// CFC twin of T_SafePulse_UserFB_Tests: the same tests drawn as CFC diagrams, the way a TwinSAFE project is authored.
    FUNCTION_BLOCK T_SafePulse_UserFB_Tests_CFC EXTENDS T_SafeCfcTestSuite
    VAR
    // Test_PulseForDelayTimeWhileInputHeld
    group_1 : T_SafeGroup;
    fb_1 : T_SafePulse_UserFB(group := group_1) := (Parameters := (DelayTime := T#100MS));
    trigStart_1 : R_TRIG;
    t1_1 : TON;
    t2_1 : TON;
    trig1_1 : R_TRIG;
    trig2_1 : R_TRIG;
    // Test_PulseEndsWhenInputDrops
    group_2 : T_SafeGroup;
    fb_2 : T_SafePulse_UserFB(group := group_2) := (Parameters := (DelayTime := T#100MS));
    // Test_StoppedGivesNoOutput
    group_3 : T_SafeGroup;
    fb_3 : T_SafePulse_UserFB(group := group_3) := (Parameters := (DelayTime := T#100MS));
    // Test_InnerBlocksJoinTheGroup
    group_4 : T_SafeGroup;
    fb_4 : T_SafePulse_UserFB(group := group_4);
END_VAR

Test_PulseForDelayTimeWhileInputHeld();
Test_PulseEndsWhenInputDrops();
Test_StoppedGivesNoOutput();
Test_InnerBlocksJoinTheGroup();

METHOD PRIVATE Test_InnerBlocksJoinTheGroup
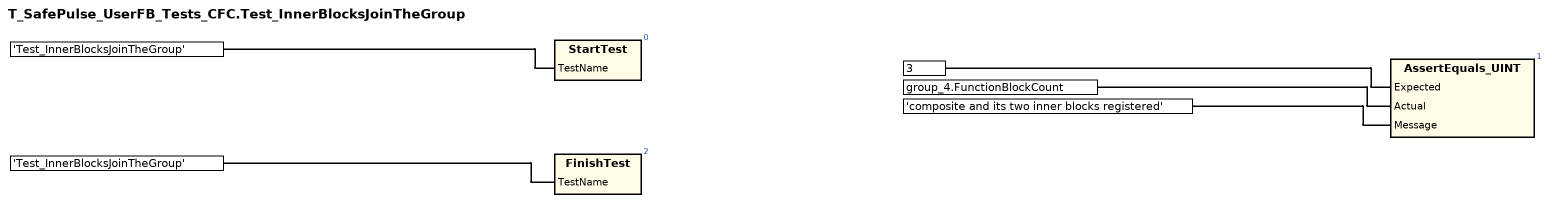
StartTest(TestName := 'Test_InnerBlocksJoinTheGroup');
AssertEquals_UINT(Expected := 3, Actual := group_4.FunctionBlockCount, Message := 'composite and its two inner blocks registered');
FinishTest(TestName := 'Test_InnerBlocksJoinTheGroup');
END_METHOD

METHOD PRIVATE Test_PulseEndsWhenInputDrops
// note: this text did not pass the execution check against the stored diagram
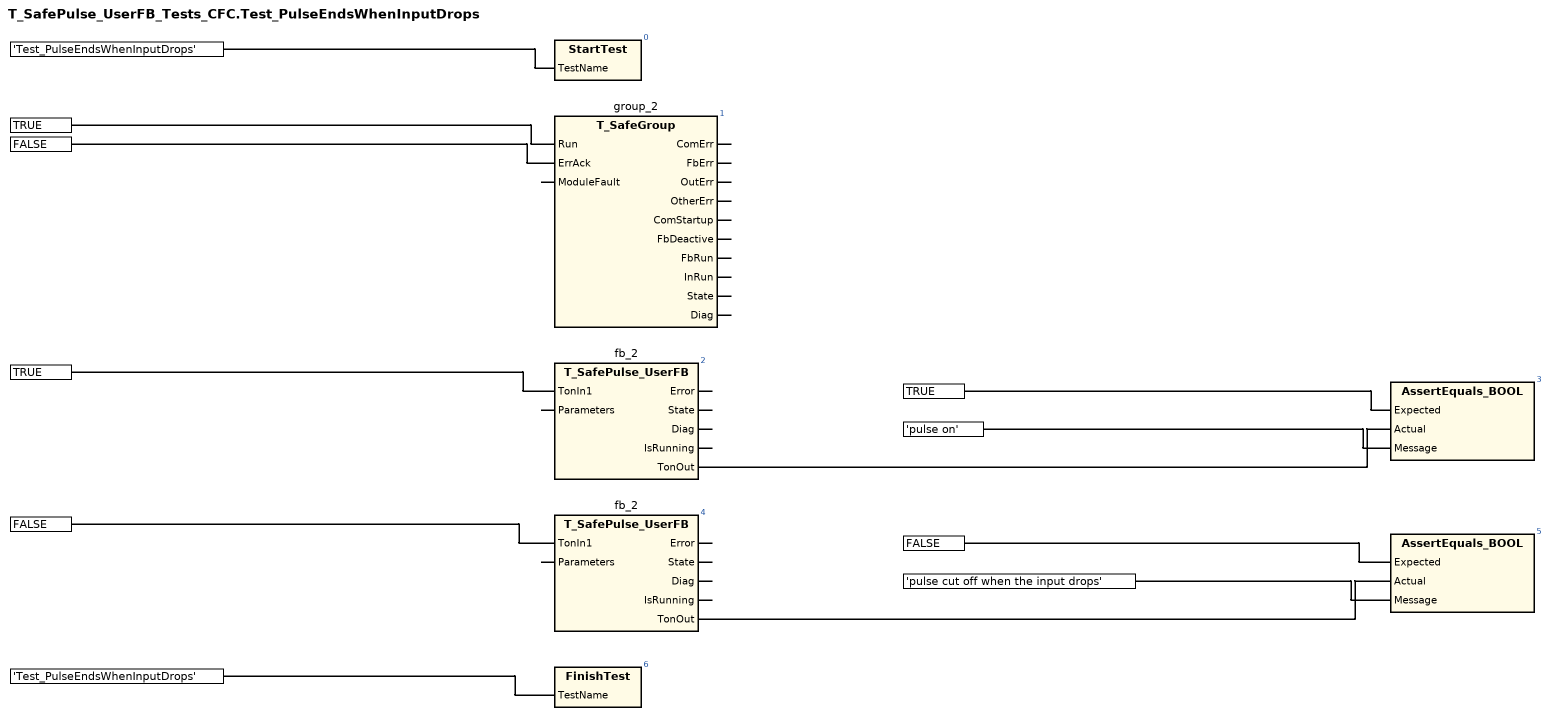
StartTest(TestName := 'Test_PulseEndsWhenInputDrops');
group_2(Run := TRUE, ErrAck := FALSE); // T_SafeGroup
fb_2(TonIn1 := TRUE); // T_SafePulse_UserFB
AssertEquals_BOOL(Expected := TRUE, Actual := fb_2.TonOut, Message := 'pulse on');
fb_2(TonIn1 := FALSE); // T_SafePulse_UserFB
AssertEquals_BOOL(Expected := FALSE, Actual := fb_2.TonOut, Message := 'pulse cut off when the input drops');
FinishTest(TestName := 'Test_PulseEndsWhenInputDrops');
END_METHOD

METHOD PRIVATE Test_PulseForDelayTimeWhileInputHeld
// note: this text did not pass the execution check against the stored diagram
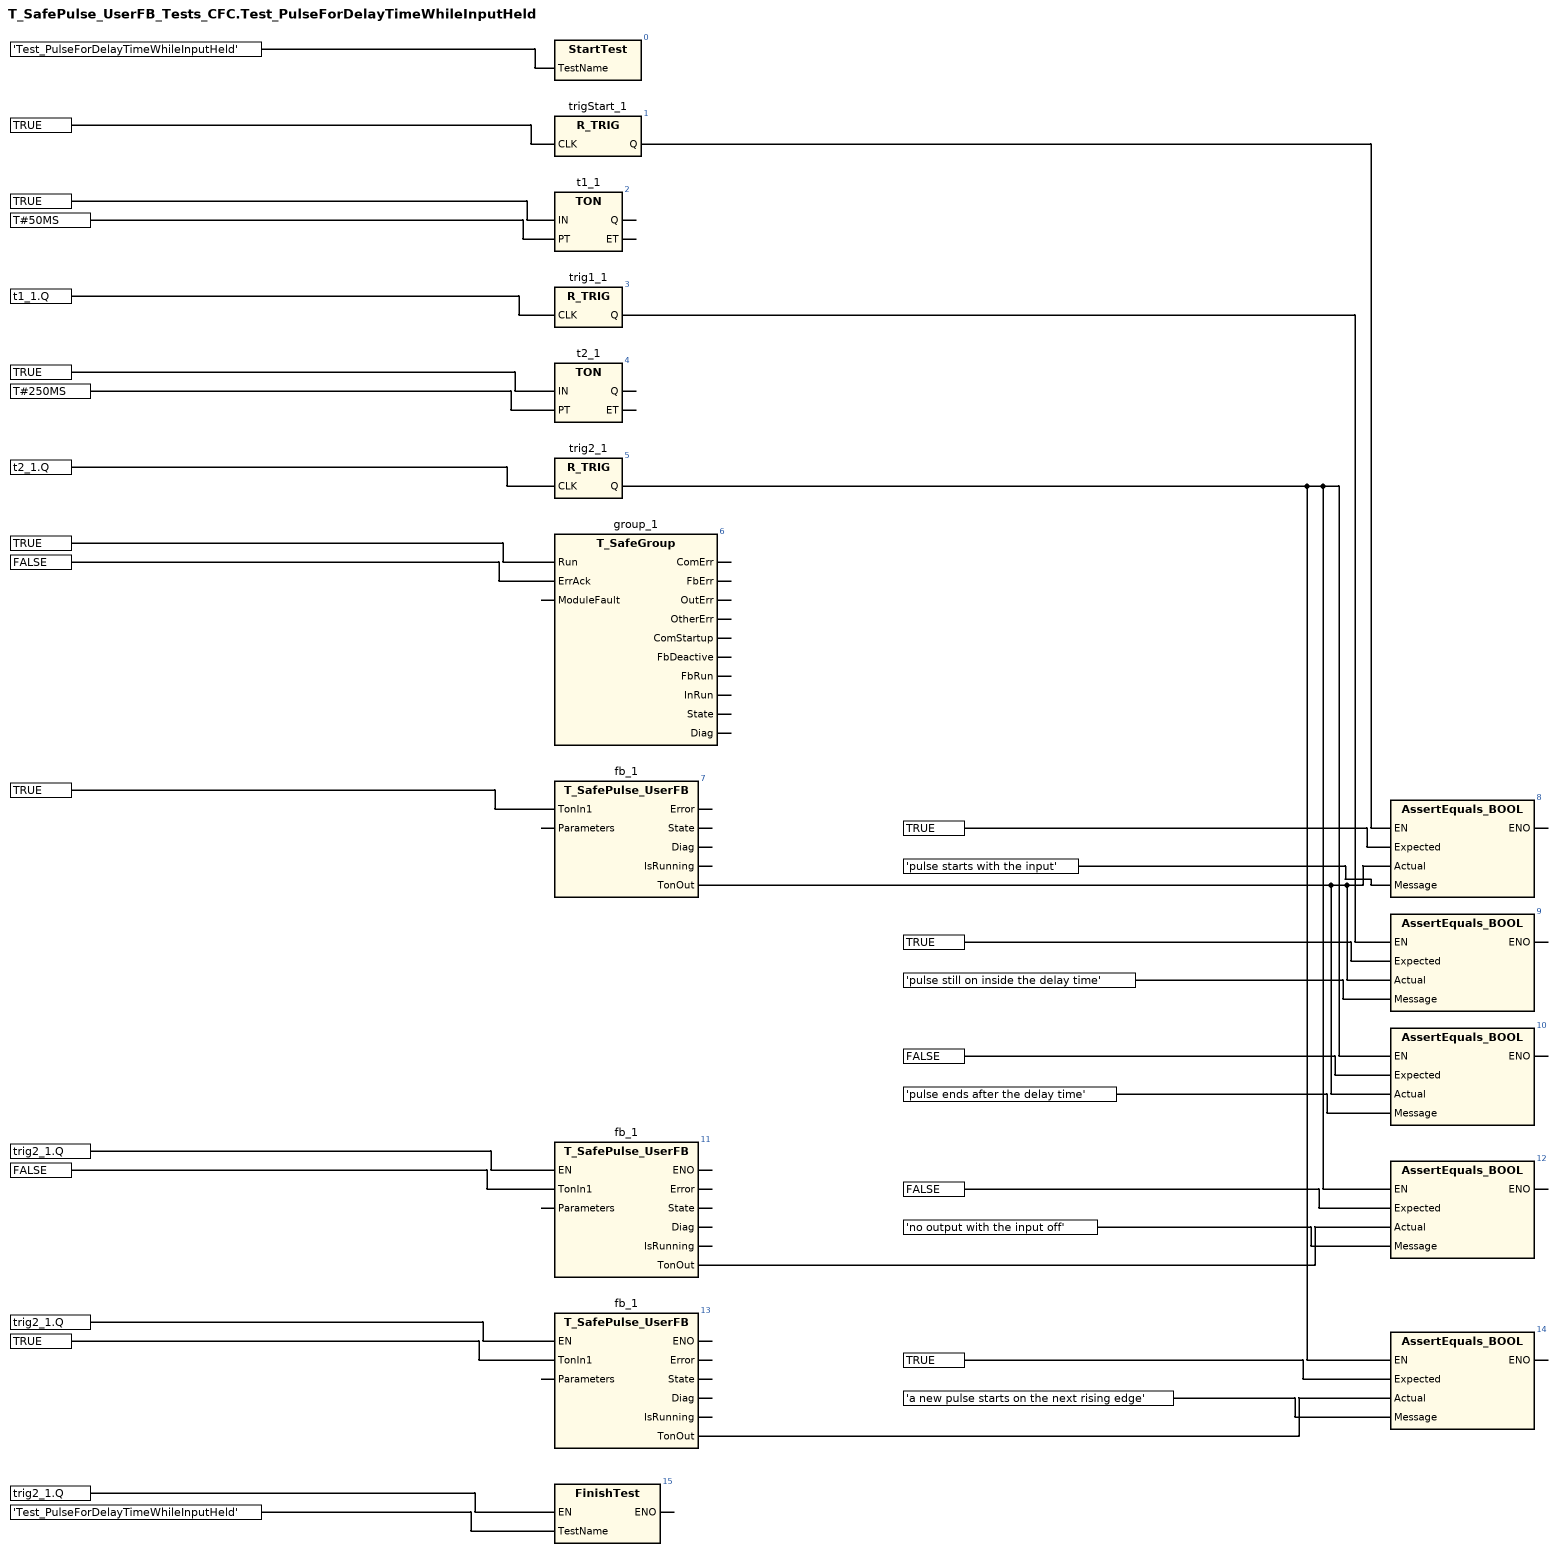
StartTest(TestName := 'Test_PulseForDelayTimeWhileInputHeld');
trigStart_1(CLK := TRUE); // R_TRIG
t1_1(IN := TRUE, PT := T#50MS); // TON
trig1_1(CLK := t1_1.Q); // R_TRIG
t2_1(IN := TRUE, PT := T#250MS); // TON
trig2_1(CLK := t2_1.Q); // R_TRIG
group_1(Run := TRUE, ErrAck := FALSE); // T_SafeGroup
fb_1(TonIn1 := TRUE); // T_SafePulse_UserFB
IF trigStart_1.Q THEN AssertEquals_BOOL(Expected := TRUE, Actual := fb_1.TonOut, Message := 'pulse starts with the input'); END_IF
IF trig1_1.Q THEN AssertEquals_BOOL(Expected := TRUE, Actual := fb_1.TonOut, Message := 'pulse still on inside the delay time'); END_IF
IF trig2_1.Q THEN AssertEquals_BOOL(Expected := FALSE, Actual := fb_1.TonOut, Message := 'pulse ends after the delay time'); END_IF
IF trig2_1.Q THEN
    fb_1(TonIn1 := FALSE); // T_SafePulse_UserFB
END_IF
IF trig2_1.Q THEN AssertEquals_BOOL(Expected := FALSE, Actual := fb_1.TonOut, Message := 'no output with the input off'); END_IF
IF trig2_1.Q THEN
    fb_1(TonIn1 := TRUE); // T_SafePulse_UserFB
END_IF
IF trig2_1.Q THEN AssertEquals_BOOL(Expected := TRUE, Actual := fb_1.TonOut, Message := 'a new pulse starts on the next rising edge'); END_IF
IF trig2_1.Q THEN FinishTest(TestName := 'Test_PulseForDelayTimeWhileInputHeld'); END_IF
END_METHOD

METHOD PRIVATE Test_StoppedGivesNoOutput
// note: this text did not pass the execution check against the stored diagram
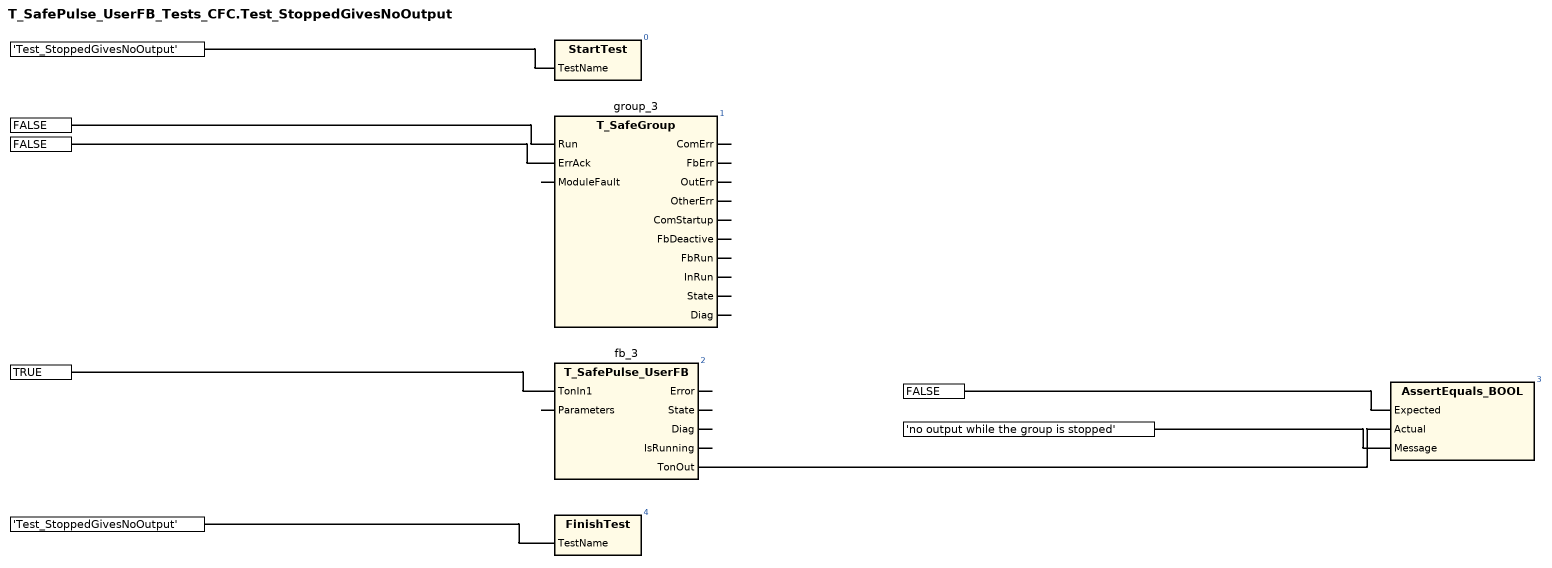
StartTest(TestName := 'Test_StoppedGivesNoOutput');
group_3(Run := FALSE, ErrAck := FALSE); // T_SafeGroup
fb_3(TonIn1 := TRUE); // T_SafePulse_UserFB
AssertEquals_BOOL(Expected := FALSE, Actual := fb_3.TonOut, Message := 'no output while the group is stopped');
FinishTest(TestName := 'Test_StoppedGivesNoOutput');
END_METHOD

END_FUNCTION_BLOCK

(* stored: Version 1.1.0.1
   POU T_SafePulse_UserFB_Tests_CFC: Id {2a8e6648-429f-5918-9f15-1d35399b8dee}, SpecialFunc None
   Method Test_InnerBlocksJoinTheGroup: Id {48313a8b-ef91-586e-bfd1-7705f670f13c}
   Method Test_PulseEndsWhenInputDrops: Id {0db4b8dc-460c-53e3-add4-566891214364}
   Method Test_PulseForDelayTimeWhileInputHeld: Id {c7a5b1db-6633-5d7f-8604-2009a54ed26d}
   Method Test_StoppedGivesNoOutput: Id {8a5f939f-b360-5360-9ec0-eacfdbbd559a} *)
